FUNCTION_BLOCK logiBUS_QDA_PWM_G (* Composite FB for 13-bit PWM output with gamma correction for lamps and LEDs (brightness 0..8191 in DWORD) *)
  (* Standard: 61499-2; Description: Copyright (c) 2026 HR Agrartechnik GmbH This program and the accompanying materials are made available under the terms of the Eclipse Public License 2.0 which is available at https://www.eclipse.org/legal/epl-2.0/ SPDX-License-Identifier: EPL-2.0 *)
  (* Version 1.0, 2026-11-06, Franz Höpfinger, HR Agrartechnik GmbH, initial version, gamma variant of logiBUS_QDA_PWM *)
  PACKAGE logiBUS::io::DQ;
  IMPORT logiBUS::io::DQ::logiBUS_DO::Invalid;
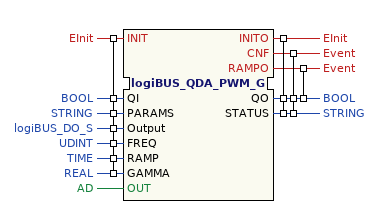
  EVENT_INPUT
    INIT : EInit WITH QI, PARAMS, Output, FREQ, RAMP, GAMMA; (* Service Initialization *)
  END_EVENT
  EVENT_OUTPUT
    INITO : EInit WITH QO, STATUS; (* Initialization Confirm *)
    CNF WITH QO, STATUS; (* Confirmation of Requested Service *)
    RAMPO WITH QO; (* Ramp finished: OUT reached (immediately after the jump with RAMP = T#0ms) *)
  END_EVENT
  VAR_INPUT
    QI : BOOL; (* Event Input Qualifier *)
    PARAMS : STRING; (* Service Parameters *)
    Output : logiBUS::io::DQ::logiBUS_DO_S := Invalid; (* Identify the Output Output_Q1..Q8 *)
    FREQ : UDINT := 400; (* PWM frequency in Hz, read at INIT. Outputs with the same frequency share an LEDC timer (4 timers, LED blinking uses one). Power stage limits, not checked: APIXON 15 PWR Q1 (BTH50030) max. 100 Hz; BTS7030/BTT6030/BTH6070 for valves 100..200 Hz; Trainer20 without power stage *)
    RAMP : TIME := T#0ms; (* Transition time to every new OUT value (hardware ramp), read at INIT. T#0ms = jump *)
    GAMMA : REAL := 2.2; (* Gamma of the brightness curve, read at INIT: duty = 8191 * (OUT / 8191)^GAMMA. 1.0 = linear (like logiBUS_QD_PWM), 2.2 = sRGB (default), 2.6 / 2.8 = Espressif examples, often more even on LEDs. Invalid values (<= 0, not finite) run linear like 1.0 *)
  END_VAR
  VAR_OUTPUT
    QO : BOOL; (* Event Output Qualifier *)
    STATUS : STRING; (* Service Status *)
  END_VAR
  SOCKETS
    OUT : adapter::types::unidirectional::AD; (* Brightness as the eye sees it (0..8191, D1), converted to the duty cycle with GAMMA *)
  END_SOCKETS
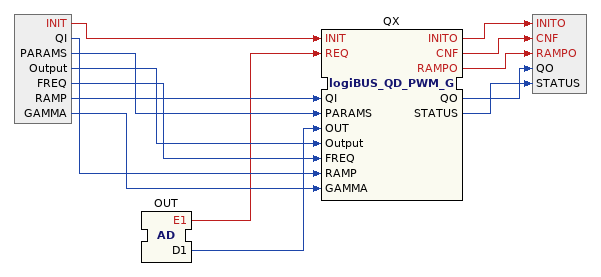
  FBS
    QX : logiBUS::io::DQ::logiBUS_QD_PWM_G;
  END_FBS
  EVENT_CONNECTIONS
    INIT TO QX.INIT;
    QX.INITO TO INITO;
    OUT.E1 TO QX.REQ;
    QX.CNF TO CNF;
    QX.RAMPO TO RAMPO;
  END_CONNECTIONS
  DATA_CONNECTIONS
    OUT.D1 TO QX.OUT;
    QI TO QX.QI;
    PARAMS TO QX.PARAMS;
    QX.QO TO QO;
    QX.STATUS TO STATUS;
    Output TO QX.Output;
    FREQ TO QX.FREQ;
    RAMP TO QX.RAMP;
    GAMMA TO QX.GAMMA;
  END_CONNECTIONS
END_FUNCTION_BLOCK
